// TIA Portal V20 export
Screen "Pop-up_AI_ENERGYMETER_Popup"  390x470
  ScreenItem "Background" at 0,0 size 390x470  Type=HmiRectangle
  ScreenItem "Textfeld_Legende" at 1,1 size 388x25  Type=HmiTextBox
  ScreenItem "Textfeld_11" at 10,33 size 285x75  Type=HmiTextBox
  ScreenItem "Textfeld_15" at 10,110 size 200x20  Type=HmiTextBox
  ScreenItem "Textfeld_16" at 10,129 size 372x71  Type=HmiTextBox
  ScreenItem "Textfeld_1" at 10,200 size 200x20  Type=HmiTextBox
  ScreenItem "Textfeld_2" at 10,220 size 372x40  Type=HmiTextBox
  ScreenItem "Textfeld_3" at 10,262 size 200x20  Type=HmiTextBox
  ScreenItem "Textfeld_4" at 10,282 size 372x20  Type=HmiTextBox
  ScreenItem "Textfeld_5" at 10,304 size 200x20  Type=HmiTextBox
  ScreenItem "Textfeld_6" at 10,324 size 372x40  Type=HmiTextBox
  ScreenItem "Textfeld_7" at 10,366 size 200x20  Type=HmiTextBox
  ScreenItem "Textfeld_8" at 10,386 size 372x20  Type=HmiTextBox
  ScreenItem "Textfeld_9" at 10,409 size 290x20  Type=HmiTextBox
  ScreenItem "Textfeld_10" at 10,427 size 372x40  Type=HmiTextBox
  ScreenItem "Cancel_Mode" at 299,1 size 90x60  Type=HmiButton
